Fanuc KAREL source: CA0106.KL

-- PROVISIONAL review KL for V770-1; original PC SHA256 3013597af57eb39015b13dc5989aba5cba3343c12ced19a3e5de8a3088317324
-- Incomplete behavior may be omitted. Consult companion uncertainty JSON. Do not deploy.
PROGRAM CA0106
%NOLOCKGROUP
BEGIN
  -- UNRESOLVED_PC offsets 0-1; opcodes 7B
  -- UNRESOLVED_PC offsets 6-22; opcodes 2D,2E,69,7F
  -- UNRESOLVED_PC offsets 27-31; opcodes 7F
  -- UNRESOLVED_PC offsets 36-43; opcodes 9C,23
  -- UNRESOLVED_PC offsets 48-55; opcodes 9D,23
  -- UNRESOLVED_PC offsets 60-71; opcodes 2E,23
  -- UNRESOLVED_PC offsets 76-83; opcodes 9D,23
  -- UNRESOLVED_PC offsets 88-97; opcodes 3F,75
  -- UNRESOLVED_PC offsets 102-116; opcodes 2E,22,9D,33,35
  -- UNRESOLVED_PC offsets 121-135; opcodes 2E,22,9D,33,35
  -- UNRESOLVED_PC offsets 140-155; opcodes 2E,22,32,35
  -- UNRESOLVED_PC offsets 160-175; opcodes 2E,22,32,35
  -- UNRESOLVED_PC offsets 180-196; opcodes 27,22,AA,23
  -- UNRESOLVED_PC offsets 201-205; opcodes 7F
END CA0106
